Fanuc KAREL source: KA00203.KL

PROGRAM KA00203
%NOLOCKGROUP
VAR
  SRC: ARRAY[4] OF VECTOR
  DST: ARRAY[4] OF BYTE
BEGIN
  DST = SRC
END KA00203
